(* IEC 61131-3 sources: genai_codesys/experiments/raw/formal/20261109_234635_2ba96d/public_02/custom__qwen3-coder-flash/attempt_01, 2 files *)

(* ---- declaration.st ---- *)
FUNCTION_BLOCK FB_DWordEdgeDetection
VAR_INPUT
    value : DWORD;
END_VAR
VAR_OUTPUT
    hasChanged : BOOL;
    hasRisingEdges : BOOL;
    risingBits : DWORD;
    noOfRisingBits : USINT;
    hasFallingEdges : BOOL;
    fallingBits : DWORD;
    noOfFallingBits : USINT;
END_VAR
VAR
    value__prev : DWORD;
END_VAR

(* ---- implementation.st ---- *)
IF value <> value__prev THEN
    hasChanged := TRUE;
ELSE
    hasChanged := FALSE;
END_IF;

risingBits := (value AND NOT value__prev);
fallingBits := (value__prev AND NOT value);

hasRisingEdges := risingBits <> 0;
hasFallingEdges := fallingBits <> 0;

noOfRisingBits := 0;
FOR i := 0 TO 31 DO
    IF (risingBits AND (1 << i)) <> 0 THEN
        noOfRisingBits := noOfRisingBits + 1;
    END_IF;
END_FOR;

noOfFallingBits := 0;
FOR i := 0 TO 31 DO
    IF (fallingBits AND (1 << i)) <> 0 THEN
        noOfFallingBits := noOfFallingBits + 1;
    END_IF;
END_FOR;

value__prev := value;
